(* IEC 61131-3 sources: llm-plc-st-eval/data/definitivo/qwen2.5-coder_14b/A4/zero_shot, 3 files *)

(* ---- ejec_1.st ---- *)
```iec
FUNCTION_BLOCK FB_Rampa
VAR_INPUT
    SPvel : REAL; // Consigna de velocidad deseada
    paroRapido : BOOL; // Indica si se debe activar el paro rápido
    ciclo : TIME; // Período de ejecución del bloque
END_VAR

VAR_OUTPUT
    CVvel : REAL; // Consigna de velocidad actual con rampa
END_VAR

VAR
    lastCVvel : REAL := 0.0; // Valor de CVvel en la última iteración
    rampaSubida : REAL := 10.0; // Pendiente de subida en puntos porcentuales por segundo
    rampaBajada : REAL := 20.0; // Pendiente de bajada en puntos porcentuales por segundo
    rampaParoRapido : REAL := 40.0; // Pendiente de paro rápido en puntos porcentuales por segundo
    tiempoCiclo : TIME := T#0s; // Tiempo transcurrido desde la última iteración
END_VAR

// Calcular el tiempo transcurrido desde la última iteración
tiempoCiclo := ciclo;

// Verificar si se debe activar el paro rápido
IF paroRapido THEN
    // Descender CVvel hacia 0.0 con la pendiente de paro rápido
    CVvel := lastCVvel - rampaParoRapido * REAL(tiempoCiclo / T#1s);
    // Asegurar que CVvel no sea menor que 0.0
    IF CVvel < 0.0 THEN
        CVvel := 0.0;
    END_IF
ELSE
    // Calcular la nueva CVvel con rampa
    IF SPvel > lastCVvel THEN
        // Subida de velocidad
        CVvel := lastCVvel + rampaSubida * REAL(tiempoCiclo / T#1s);
        // Asegurar que CVvel no supere el valor objetivo
        IF CVvel > SPvel THEN
            CVvel := SPvel;
        END_IF
    ELSE
        // Bajada de velocidad
        CVvel := lastCVvel - rampaBajada * REAL(tiempoCiclo / T#1s);
        // Asegurar que CVvel no sea menor que el valor objetivo
        IF CVvel < SPvel THEN
            CVvel := SPvel;
        END_IF
    END_IF
END_IF

// Actualizar el valor de lastCVvel para la próxima iteración
lastCVvel := CVvel;
END_FUNCTION_BLOCK
```

(* ---- ejec_2.st ---- *)
```pascal
FUNCTION_BLOCK FB_Rampa
VAR_INPUT
    SPvel : REAL;       // Consigna de velocidad deseada
    paroRapido : BOOL;  // Indica si se debe activar el paro rápido
    ciclo : TIME;       // Período de ejecución del bloque
END_VAR

VAR_OUTPUT
    CVvel : REAL;       // Consigna de velocidad actual
END_VAR

VAR
    lastCVvel : REAL;   // Valor de CVvel en la iteración anterior
    rampaSubida : REAL := 10.0;  // Pendiente de subida en puntos porcentuales por segundo
    rampaBajada : REAL := 20.0;  // Pendiente de bajada en puntos porcentuales por segundo
    rampaParoRapido : REAL := 40.0;  // Pendiente de paro rápido en puntos porcentuales por segundo
    tiempoCiclo : TIME;  // Tiempo transcurrido desde la última iteración
END_VAR

// Calcular el tiempo transcurrido desde la última iteración
tiempoCiclo := ciclo;

// Verificar si se debe activar el paro rápido
IF paroRapido THEN
    // Descender CVvel hacia 0.0 con una pendiente de 40.0 puntos porcentuales por segundo
    CVvel := MAX(0.0, lastCVvel - rampaParoRapido * REAL(tiempoCiclo / T#1s));
ELSE
    // Calcular la nueva CVvel según la consigna SPvel
    IF SPvel > lastCVvel THEN
        // Subida de velocidad
        CVvel := MIN(SPvel, lastCVvel + rampaSubida * REAL(tiempoCiclo / T#1s));
    ELSE
        // Bajada de velocidad
        CVvel := MAX(SPvel, lastCVvel - rampaBajada * REAL(tiempoCiclo / T#1s));
    END_IF;
END_IF;

// Actualizar el valor de lastCVvel para la próxima iteración
lastCVvel := CVvel;
```

Este código implementa un generador de consigna de velocidad con rampa en un FUNCTION_BLOCK llamado `FB_Rampa`. La salida `CVvel` sigue a la consigna `SPvel` con las pendientes especificadas, y en caso de activación de `paroRapido`, `CVvel` descenderá hacia 0.0 con una pendiente de 40.0 puntos porcentuales por segundo.

(* ---- ejec_3.st ---- *)
```iec
FUNCTION_BLOCK FB_Rampa
VAR_INPUT
    SPvel : REAL; // Consigna de velocidad deseada
    paroRapido : BOOL; // Indicador de paro rápido
    ciclo : TIME; // Período de ejecución del bloque
END_VAR

VAR_OUTPUT
    CVvel : REAL; // Consigna de velocidad actualizada con rampa
END_VAR

VAR
    error : REAL; // Diferencia entre SPvel y CVvel
    deltaCVvel : REAL; // Cambio en CVvel durante el ciclo
    maxRampaSubida : REAL := 10.0; // Máxima rampa de subida en puntos porcentuales por segundo
    maxRampaBajada : REAL := 20.0; // Máxima rampa de bajada en puntos porcentuales por segundo
    maxRampaParoRapido : REAL := 40.0; // Máxima rampa de paro rápido en puntos porcentuales por segundo
    cicloSegundos : REAL; // Ciclo convertido a segundos
END_VAR

// Convertir el ciclo de tiempo a segundos
cicloSegundos := REAL(ciclo) / 1000.0;

// Calcular el error entre la consigna deseada y la actual
error := SPvel - CVvel;

// Determinar el cambio en CVvel según las condiciones
IF paroRapido THEN
    // Modo paro rápido: descender hacia 0 con una pendiente máxima
    deltaCVvel := -maxRampaParoRapido * cicloSegundos;
    IF CVvel + deltaCVvel < 0.0 THEN
        CVvel := 0.0;
    ELSE
        CVvel := CVvel + deltaCVvel;
    END_IF
ELSE
    // Modo normal: seguir la consigna con rampa
    IF error > 0 THEN
        // Subida de velocidad
        deltaCVvel := maxRampaSubida * cicloSegundos;
        IF CVvel + deltaCVvel > SPvel THEN
            CVvel := SPvel;
        ELSE
            CVvel := CVvel + deltaCVvel;
        END_IF
    ELSE
        // Bajada de velocidad
        deltaCVvel := -maxRampaBajada * cicloSegundos;
        IF CVvel + deltaCVvel < SPvel THEN
            CVvel := SPvel;
        ELSE
            CVvel := CVvel + deltaCVvel;
        END_IF
    END_IF
END_IF;

END_FUNCTION_BLOCK
```
